Fanuc KAREL source: ka00165.KL

PROGRAM KA00165
%STACKSIZE=65535
%PRIORITY=65535
%NOLOCKGROUP
VAR
SRC : ARRAY[4] OF BOOLEAN
DST : ARRAY[4] OF BOOLEAN
BEGIN
-- UNRESOLVED_PC line 7 opcodes [22 22 1E] marker_code=0
END KA00165
